(* PLC project Vn_fanout_two_wires, Beckhoff Automation GmbH TwinCAT PLC Control 3.5.13.21 *)
(* stored: creationDateTime 1970-01-01T00:00:00 *)

PROGRAM Vn_fanout_two_wires
  VAR  (* added by the conversion: wires and edge detectors of the diagram *)
    _AND10000000003_OUT : BOOL;
    _OR10000000006_OUT : BOOL;
  END_VAR

(* FBD diagram, written out as Structured Text *)
_AND10000000003_OUT := a AND b;
_OR10000000006_OUT := c OR d;
out1 := _AND10000000003_OUT AND _OR10000000006_OUT;
out2 := _AND10000000003_OUT OR _OR10000000006_OUT;
END_PROGRAM
